INTERFACE I_Alarm EXTENDS I_CatalogEvent

METHOD Raise : HRESULT
END_METHOD

METHOD Clear : HRESULT
VAR_INPUT
	bResetConfirmation	: BOOL;
END_VAR
END_METHOD

METHOD Confirm : HRESULT
END_METHOD

// Level driven: raises while bActive is TRUE, clears when it drops.
METHOD SetActive : HRESULT
VAR_INPUT
	bActive	: BOOL;
END_VAR
END_METHOD

PROPERTY IsRaised : BOOL
GET
END_GET
END_PROPERTY

PROPERTY ConfirmationState : TcEventConfirmationState
GET
END_GET
END_PROPERTY

END_INTERFACE

(* stored: Version 1.1.0.1, ProductVersion 3.1.4026.26
   Itf I_Alarm: Id {4bfdbc82-0539-4d6a-8ea5-737cf605239b}
   Method Raise: Id {e5a91d98-6862-4ddd-9c37-2efdb32df127}
   Method Clear: Id {a0763371-6747-44f4-8bf6-354d8f22101a}
   Method Confirm: Id {d613ac01-ac15-48ad-b6bc-a4a568bb8915}
   Method SetActive: Id {477af543-31aa-4bf3-9506-0c6d4601fa71}
   Property IsRaised: Id {28937878-11ef-4f0b-abe0-0f149e093da2}
   Get Get: Id {ccf2ba70-be33-4889-bdcc-62561fd267ea}
   Property ConfirmationState: Id {15f50921-164f-4c46-8eee-5b06bdd1353d}
   Get Get: Id {bcc5249d-e193-4429-8bd5-3eeb0c193189} *)
